(* IEC 61131-3 sources: plcassist-cli/packages/volt-lsp-iec/test-corpus/awa-palletizer/Device/Plc Logic/Application/Library Manager/(unresolved)/cmpeventmgr interfaces, 3 files *)

(* ---- CONSTANTS.gvl ---- *)
VAR_GLOBAL
	EVENT_CALLBACKS_NO_LIMIT : UDINT := 16#FFFFFFFF;
	CMPID_CMPEVENTMGR : UDINT := 16#5B;
	ITFID_ICMPEVENTCALLBACK : UDINT := 16#25;
END_VAR

(* ---- EVENTCLASS.gvl ---- *)
VAR_GLOBAL
	EVTCLASS_NONE : UINT := 0;
	EVTCLASS_ALL : UINT := 16#FFFF;
	EVTCLASS_INFO : UINT := 16#1;
	EVTCLASS_WARNING : UINT := 16#2;
	EVTCLASS_ERROR : UINT := 16#4;
	EVTCLASS_EXCEPTION : UINT := 16#8;
	EVTCLASS_VENDOR_SPEC : UINT := 16#1000;
END_VAR

(* ---- ICMPEVENTCALLBACK.itf ---- *)
INTERFACE ICMPEVENTCALLBACK
END_INTERFACE

METHOD EVENTCALLBACK : RTS_IEC_RESULT
VAR_INPUT
	PEVENTPARAM : POINTER TO EventParam;
END_VAR
END_METHOD
